Fanuc KAREL source: kt00747.KL

PROGRAM KT00747
%STACKSIZE=65535
%PRIORITY=65535
%NOLOCKGROUP
VAR
ARG : ARRAY[4] OF JOINTPOS9
OUT : INTEGER
BEGIN
-- UNSAFE_SOURCE_IR line 7: OUT = native_s16_value(ARG)
END KT00747
